{attribute 'pack_mode' := '2'}
TYPE ST_INSTANCE_STATE :
STRUCT
  ProcessIdentity   : E_INSTANCE;

  ProcessState      : E_INSTANCE_STATE;
  ProcessProgress   : E_PROGRESS;

  CollectorState    : E_PROCESS_STATE;
  CollectorProgress : E_PROGRESS;
  CollectorCheck    : E_PROCESS_CHECK;

  QueueProcessCount : UINT; // sum of all queues in process
  StationCount      : UINT;
  ListCount         : UINT; // number of tickets in ProcessList
END_STRUCT
END_TYPE

(* stored: Version 1.1.0.1
   DUT ST_INSTANCE_STATE: Id {7108ed74-ad9f-421c-8515-268b082913f8} *)
